(* IEC 61131-3 sources: Gen-AI/final/Gen-AI_v1.0_submission/A2_框架源码/agent/logs/full34_fixture/E3_S14_1_42/tools/candidate_1/fixture_compile, 1 file *)

(* ---- source.st ---- *)
FUNCTION_BLOCK FB_S14
VAR_INPUT
    Pressure : REAL;
    PumpEnable : BOOL;
    ResetBtn : BOOL;
END_VAR
VAR_OUTPUT
    LowPump : BOOL;
    HighPump : BOOL;
    ReliefValve : BOOL;
    AlarmLamp : BOOL;
    Status : WORD;
END_VAR
(* Add a VAR block for internal state/timers before the implementation, if needed. *)
(* SKELETON ONLY: replace this RETURN with scan logic and required initial state. *)
RETURN;
END_FUNCTION_BLOCK

(* FIXTURE_COMPILE_FAIL *)
